(* IEC 61131-3 sources: plcassist-cli/packages/volt-lsp-iec/test-corpus/pro2193/Device/Plc Logic/Application/09 Misc/Library Manager/(unresolved)/base interfaces, 3 files *)

(* ---- COMPONENTIDS.gvl ---- *)
VAR_GLOBAL
	CMPID_IECCODE : DWORD := 16#1000;
	CMPID_CMPSTARTOEM : DWORD := 16#2000;
	CMPID_CMPENDOEM : DWORD := 16#3FFF;
END_VAR

(* ---- INTERFACEIDS.gvl ---- *)
VAR_GLOBAL
	ITFID_IBASE : DWORD := 16#0;
	ITFID_ICMPSTARTOEM : DWORD := 16#2000;
	ITFID_ICMPENDOEM : DWORD := 16#3FFF;
END_VAR

(* ---- IBASE.itf ---- *)
INTERFACE IBASE
END_INTERFACE

METHOD FB_EXIT : BOOL
VAR_INPUT
	BINCOPYCODE : BOOL;
END_VAR
END_METHOD

METHOD RELEASE : DINT
END_METHOD

METHOD FB_REINIT : BOOL
END_METHOD

METHOD ADDREF : DINT
END_METHOD

METHOD QUERYINTERFACE : POINTER TO POINTER TO BYTE
VAR_INPUT
	IID : DWORD;
	PRESULT : POINTER TO UDINT;
END_VAR
END_METHOD

METHOD FB_INIT : BOOL
VAR_INPUT
	BINITRETAINS : BOOL;
	BINCOPYCODE : BOOL;
END_VAR
END_METHOD
